(* IEC 61131-3 sources: model-first-plc-agent-ai/results/T2-B-22, 1 file *)

(* ---- b_code.st ---- *)
FUNCTION_BLOCK FillingControl
VAR_INPUT
    start : BOOL;
    stop : BOOL;
    LSH : BOOL;
    LSHH : BOOL;
    TimerDuration : TIME;
END_VAR
VAR_OUTPUT
    fill_valve : BOOL;
    discharge_valve : BOOL;
END_VAR
VAR
    current_state : INT := 0;
    filling_timer : TON;
    timer_done : BOOL := FALSE;
END_VAR

(* Stop has priority. High-high level prevents or terminates filling. *)
IF stop OR LSHH THEN
    current_state := 0;
ELSE
    CASE current_state OF
        0:
            IF start THEN
                current_state := 1;
            END_IF;
        1:
            current_state := 1;
    ELSE
        current_state := 0;
    END_CASE;
END_IF;

filling_timer(
    IN := (current_state = 1),
    PT := TimerDuration
);
timer_done := filling_timer.Q;

IF (current_state = 1) AND timer_done THEN
    current_state := 0;
    (* Reset immediately so a later start always gets a fresh interval. *)
    filling_timer(IN := FALSE, PT := TimerDuration);
END_IF;

fill_valve := (current_state = 1) AND NOT stop AND NOT LSHH;
discharge_valve := FALSE;

END_FUNCTION_BLOCK

PROGRAM Main
VAR
    StartCommand AT %IX100.0 : BOOL;
    StopCommand AT %IX100.1 : BOOL;
    LSH AT %IX100.2 : BOOL;
    LSHH AT %IX100.3 : BOOL;
    FillValve AT %QX100.0 : BOOL;
    DischargeValve AT %QX100.1 : BOOL;
END_VAR
VAR
    (* Configurable filling interval. *)
    TimerDuration : TIME := T#10s;
    start_edge : R_TRIG;
    controller : FillingControl;
END_VAR

start_edge(CLK := StartCommand);

controller(
    start := start_edge.Q,
    stop := StopCommand,
    LSH := LSH,
    LSHH := LSHH,
    TimerDuration := TimerDuration
);

FillValve := controller.fill_valve;
DischargeValve := controller.discharge_valve;

END_PROGRAM
